(* CODESYS project AddJobDialog.xml

Project tree, tasks and I/O mapping:
  visualisation AddJobDialog
*)

// /AddJobDialog
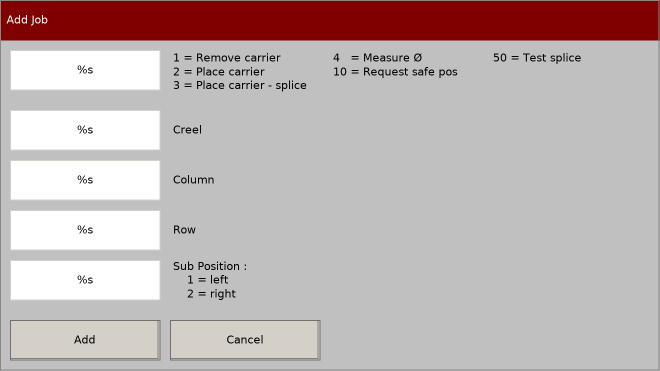
VISUALIZATION AddJobDialog  // 660x371
    Rectangle (0,40 660x331)
    Label (170,110 150x40), "Creel"
    Label (170,210 150x40), "Row"
    Label (170,260 150x40), "Sub Position : 1 = left 2 = right"
    Textfield (10,110 150x40), "%s", text variable: PRG_VisuTask_10ms._fbJobMgrCtrl._scCreelPos.scCreelPos.eCreel
        OnMouseUp: write the text variable via Default
    Textfield (10,210 150x40), "%s", text variable: PRG_VisuTask_10ms._fbJobMgrCtrl._scCreelPos.scCreelPos.uiRow
        OnMouseUp: write the text variable via Default
    Textfield (10,260 150x40), "%s", text variable: PRG_VisuTask_10ms._fbJobMgrCtrl._scCreelPos.scCreelPos.eSubPosition
        OnMouseUp: write the text variable via Default
    Rectangle (170,50 150x40), "1 = Remove carrier 2 = Place carrier 3 = Place carrier - splice"
    Textfield (10,50 150x40), "%s", text variable: PRG_VisuTask_10ms._fbJobMgrCtrl._scCreelPos.eType
        OnMouseUp: write the text variable via Default
    Rectangle (330,50 150x40), "4 = Measure Ø 10 = Request safe pos"
    Button (10,320 150x40), "Add"
        tap PRG_VisuTask_10ms._fbJobMgrCtrl._btnAddJob.xbtn
        OnMouseUp:  Dialog=AddJobDialog, Result=OK, NumpadKeypadSet=True
    Button (170,320 150x40), "Cancel"
        OnMouseUp:  Dialog=AddJobDialog, Result=OK, NumpadKeypadSet=True
    Rectangle (0,0 660x40), "Add Job"
    Rectangle (490,50 150x40), "50 = Test splice"
    Label (170,160 150x40), "Column"
    Textfield (10,160 150x40), "%s", text variable: PRG_VisuTask_10ms._fbJobMgrCtrl._scCreelPos.scCreelPos.uiColumn
        OnMouseUp: write the text variable via Default
END_VISUALIZATION
